(* IEC 61131-3 sources: volt/packages/volt-lsp-iec/test-corpus/pro2193/Device/Plc Logic/Application/09 Misc/Library Manager/L_IOM_IOModules, 22 files *)

(* ---- L_IOM_FAST_OUTP.dut ---- *)
TYPE L_IOM_FAST_OUTP :
STRUCT
	BYVALUE : BYTE;
	BYRUNNINGNUMBER : BYTE;
	WTIMETICK : WORD;
	DWTIMETICK : DWORD;
	XINUSE : BOOL;
END_STRUCT
END_TYPE

(* ---- L_IOM_FAST_OUTP_UNSORTED.dut ---- *)
TYPE L_IOM_FAST_OUTP_UNSORTED :
STRUCT
	BYDIGITALOUTPUTSEL : BYTE;
	BYVALUE : BYTE;
	WTIMETICK : WORD;
	DWTIMETICK : DWORD;
	XINUSE : BOOL;
END_STRUCT
END_TYPE

(* ---- L_IOM_FAST_RXTXPDO.dut ---- *)
TYPE L_IOM_FAST_RXTXPDO :
STRUCT
	WNUMBEROFEXCLUDES : WORD;
	WNUMBEROFENTRIES : WORD;
	WINDEX : WORD;
	BYFIXED : BYTE;
	BYMANDATORY : BYTE;
	WVIRTUAL : WORD;
	WSM : WORD;
	WSU : WORD;
	SNAME : STRING;
END_STRUCT
END_TYPE

(* ---- L_IOM_FAST_TXPDO.dut ---- *)
TYPE L_IOM_FAST_TXPDO :
STRUCT
	WINDEX : WORD;
	WSUBINDEX : WORD;
	WSIZE : WORD;
END_STRUCT
END_TYPE

(* ---- L_IOM_FASTIO_IO_ADDRESSES.dut ---- *)
TYPE L_IOM_FASTIO_IO_ADDRESSES :
STRUCT
	PBYVALUE : POINTER TO BYTE;
	PBYRUNNINGNUMBER : POINTER TO BYTE;
	PWTIMETICK : POINTER TO WORD;
END_STRUCT
END_TYPE

(* ---- L_IOM_FASTIO_OUT_STATE_INPUT.dut ---- *)
TYPE L_IOM_FASTIO_OUT_STATE_INPUT :
STRUCT
	PBYLASTRUNNINGNUMBER : POINTER TO BYTE;
	PBYNEXTRUNNINGNUMBER : POINTER TO BYTE;
	PBYSTATEFIFO : POINTER TO BYTE;
	PBYCOUNTFIFOENTRIES : POINTER TO BYTE;
	PDWABSOLUTECOUNTER : POINTER TO DWORD;
END_STRUCT
END_TYPE

(* ---- L_IOM_IEXTERNALTPINTERFACE.itf ---- *)
INTERFACE L_IOM_IEXTERNALTPINTERFACE
END_INTERFACE

METHOD CHECKABORTED : BOOL
VAR_INPUT
	TOUCHPROBECHANNEL : BYTE;
END_VAR
END_METHOD

METHOD CHECKCONFIGURATION : BOOL
VAR_INPUT
	TOUCHPROBESOURCE : BYTE;
	TOUCHPROBECHANNEL : BYTE;
	TOUCHPROBESIGNAL : BYTE;
	TOUCHPROBEEDGE : BYTE;
	TOUCHPROBEMODE : BYTE;
END_VAR
VAR_OUTPUT
	WERRORID : WORD := 0;
END_VAR
END_METHOD

METHOD CHECKNEWTP : BOOL
VAR_INPUT
	TOUCHPROBECHANNEL : BYTE;
	TOUCHPROBEEDGE : BYTE;
END_VAR
VAR_OUTPUT
	XTPPOSEDGE : BOOL;
	XTPNEGEDGE : BOOL;
	WTPTIMETICKPOSEDGE : WORD;
	WTPTIMETICKNEGEDGE : WORD;
	DWTPTIMETICKABSCOUNTER : DWORD;
END_VAR
END_METHOD

METHOD INITFORNEWTP : BOOL
VAR_INPUT
	TOUCHPROBECHANNEL : BYTE;
END_VAR
END_METHOD

METHOD SETABORT : BOOL
VAR_INPUT
	TOUCHPROBECHANNEL : BYTE;
END_VAR
END_METHOD

(* ---- CALCRXPDOOFFSETS131.pou ---- *)
FUNCTION CALCRXPDOOFFSETS131 : BOOL
VAR_INPUT
	PCONNECTOR : POINTER TO IoConfigConnector;
	WSLICEPOSITION : WORD;
	WPDOOFFSETBASE : WORD;
END_VAR
VAR_OUTPUT
	WPDOOFFSET : WORD;
	WPDONUMBEROFENTRIES : WORD;
END_VAR
END_FUNCTION

(* ---- CALCTXPDOOFFSETS131.pou ---- *)
FUNCTION CALCTXPDOOFFSETS131 : BOOL
VAR_INPUT
	PCONNECTOR : POINTER TO IoConfigConnector;
	WSLICEPOSITION : WORD;
	WPDOOFFSETBASE : WORD;
END_VAR
VAR_OUTPUT
	WPDOOFFSET : WORD;
	WPDONUMBEROFENTRIES : WORD;
END_VAR
END_FUNCTION

(* ---- FINDOWNSLICEPOSITIONS131.pou ---- *)
FUNCTION FINDOWNSLICEPOSITIONS131 : BOOL
VAR_INPUT
	M_HINTERFACE : POINTER TO IoConfigConnector;
	M_PCONNECTOR : POINTER TO IoConfigConnector;
	WMODULETYPE : WORD;
END_VAR
VAR_OUTPUT
	WSLICEPOSITION : WORD;
END_VAR
END_FUNCTION

(* ---- GETBOOLEANPROPERTY.pou ---- *)
FUNCTION GETBOOLEANPROPERTY : BOOL
VAR_INPUT
	STKEY : WSTRING;
END_VAR
END_FUNCTION

(* ---- GETCOMPANY.pou ---- *)
FUNCTION GETCOMPANY : WSTRING
END_FUNCTION

(* ---- GETNUMBERPROPERTY.pou ---- *)
FUNCTION GETNUMBERPROPERTY : DINT
VAR_INPUT
	STKEY : WSTRING;
END_VAR
END_FUNCTION

(* ---- GETTEXTPROPERTY.pou ---- *)
FUNCTION GETTEXTPROPERTY : WSTRING
VAR_INPUT
	STKEY : WSTRING;
END_VAR
END_FUNCTION

(* ---- GETTEXTPROPERTY2.pou ---- *)
FUNCTION GETTEXTPROPERTY2 : POINTER TO WSTRING
VAR_INPUT
	STKEY : WSTRING;
END_VAR
END_FUNCTION

(* ---- GETTITLE.pou ---- *)
FUNCTION GETTITLE : WSTRING
END_FUNCTION

(* ---- GETVERSION.pou ---- *)
FUNCTION GETVERSION : VERSION
END_FUNCTION

(* ---- GETVERSIONPROPERTY.pou ---- *)
FUNCTION GETVERSIONPROPERTY : VERSION
VAR_INPUT
	STKEY : WSTRING;
END_VAR
END_FUNCTION

(* ---- L_FASTIO_INREF.pou ---- *)
FUNCTION_BLOCK L_FASTIO_INREF EXTENDS IoDrvBase
VAR_INPUT
	XAABORTISACTIVE : ARRAY [0..3] OF BOOL;
END_VAR
VAR_OUTPUT
	IOVARIABLEADDRESSES : ARRAY [0..(FIFO_SIZE_MAX - 1)] OF L_IOM_FASTIO_IO_ADDRESSES;
	BYRISINGEDGEPARAMETERVALUE : BYTE;
	BYFALLINGEDGEPARAMETERVALUE : BYTE;
	BYMAXTPCOUNT : BYTE := 2;
	PDWABSOLUTECOUNTER : POINTER TO DWORD;
END_VAR
VAR
	CMPID_CMPLENZEFASTIO_INREF : DWORD := 16#1028200B;
	FIFO_SIZE_MAX : BYTE := 15;
	PARAM_ID_MODUL_IDENT : DWORD := 16#41000000;
	MODUL_IDENT_S207 : DWORD := 16#F0147C1;
	MODUL_IDENT_S208 : DWORD := 16#F0347C2;
	M_IIODRV : ICmpIoDrv;
	M_IIODRVPARAMETER : ICmpIoDrvParameter;
	XINPUTSVALID : BOOL := TRUE;
	XINPUTSVALIDACTCYCLE : BOOL := TRUE;
	XFIRSTEDGEDETECTED : BOOL := FALSE;
	ILASTRUNNINGNUMBER : ARRAY [1..4] OF INT := [-1, -1, -1, -1];
	BYNEWSIGNAL : ARRAY [1..4] OF BYTE := [0, 0, 0, 0];
	BYOLDSIGNAL : ARRAY [1..4] OF BYTE := [0, 0, 0, 0];
	FIFO_SIZE : BYTE;
	PMYFATHERCONNECT_68 : POINTER TO IoConfigConnector;
	PMYGRANDFATHERCONNECT_65 : POINTER TO IoConfigConnector;
	DWMODULIDENT : DWORD;
	PRESULT : POINTER TO SysTypes.RTS_IEC_RESULT;
	_XINITIALINPUTSTATEAVAILABLE : BOOL := FALSE;
	_ABYINITIALINPUTSTATE : ARRAY [0..1] OF BYTE;
	XFIRSTEDGETIMESTAMPVALID : BOOL := FALSE;
	DWFIRSTEDGETIMESTAMP : DWORD;
	BYINITIALINPUTSTATE : BYTE;
	FIRSTEDGEDETECTED : BOOL;
END_VAR
END_FUNCTION_BLOCK

METHOD INITIALIZE : UDINT
VAR_INPUT
	WMODULETYPE : UINT;
	DWINSTANCE : UDINT;
	PCONNECTOR : POINTER TO IoConfigConnector;
END_VAR
END_METHOD

METHOD FB_INIT : BOOL
VAR_INPUT
	BINITRETAINS : BOOL;
	BINCOPYCODE : BOOL;
END_VAR
END_METHOD

METHOD QUERYINTERFACE : POINTER TO POINTER TO BYTE
VAR_INPUT
	IID : DWORD;
	PRESULT : POINTER TO UDINT;
END_VAR
END_METHOD

METHOD IODRVUPDATECONFIGURATION : UDINT
VAR_INPUT
	PCONNECTORLIST : POINTER TO IoConfigConnector;
	NCOUNT : DINT;
END_VAR
END_METHOD

METHOD IODRVUPDATEMAPPING : UDINT
VAR_INPUT
	PTASKMAPLIST : POINTER TO IoConfigTaskMap;
	NCOUNT : DINT;
END_VAR
END_METHOD

METHOD IODRVGETCONNECTOR : POINTER TO IoConfigConnector
VAR_INPUT
	PRESULT : POINTER TO SysTypes.RTS_IEC_RESULT;
END_VAR
END_METHOD

METHOD CHECKABORTED : BOOL
VAR_INPUT
	TOUCHPROBECHANNEL : BYTE;
END_VAR
END_METHOD

METHOD CHECKCONFIGURATION : BOOL
VAR_INPUT
	TOUCHPROBESOURCE : BYTE;
	TOUCHPROBECHANNEL : BYTE;
	TOUCHPROBESIGNAL : BYTE;
	TOUCHPROBEEDGE : BYTE;
	TOUCHPROBEMODE : BYTE;
END_VAR
VAR_OUTPUT
	WERRORID : WORD := 0;
END_VAR
END_METHOD

METHOD CHECKNEWTP : BOOL
VAR_INPUT
	TOUCHPROBECHANNEL : BYTE;
	TOUCHPROBEEDGE : BYTE;
END_VAR
VAR_OUTPUT
	XTPPOSEDGE : BOOL;
	XTPNEGEDGE : BOOL;
	WTPTIMETICKPOSEDGE : WORD;
	WTPTIMETICKNEGEDGE : WORD;
	DWTPTIMETICKABSCOUNTER : DWORD;
END_VAR
END_METHOD

METHOD EDGEDETECTED : BOOL
VAR_INPUT
	TOUCHPROBEEDGE : BYTE;
	BYNEWSIGNAL : BYTE;
	BYOLDSIGNAL : BYTE;
	WTIMETICK : WORD;
END_VAR
VAR_OUTPUT
	XTPPOSEDGE : BOOL;
	XTPNEGEDGE : BOOL;
	WTPTIMETICKPOSEDGE : WORD;
	WTPTIMETICKNEGEDGE : WORD;
END_VAR
END_METHOD

METHOD INITFORNEWTP : BOOL
VAR_INPUT
	TOUCHPROBECHANNEL : BYTE;
END_VAR
END_METHOD

METHOD SETABORT : BOOL
VAR_INPUT
	TOUCHPROBECHANNEL : BYTE;
END_VAR
END_METHOD

(* ---- L_FASTIO_INREF_ECAT.pou ---- *)
FUNCTION_BLOCK L_FASTIO_INREF_ECAT EXTENDS L_FastIO_InRef
VAR
	WINITSTATE : WORD := 0;
	DWBUFFER : DWORD;
	L_ETC_COE_SDOWRITE1 : L_ETC_CoE_SdoWrite;
	L_ETC_GETMASTERSTATE1 : L_ETC_GetMasterState;
	WSLICEPOSITION : WORD;
	WPDOOFFSET : WORD;
	WPDONUMBEROFENTRIES : WORD;
	WECATSLAVEADR : WORD;
	PDWABSOLUTECOUNTERBPB : POINTER TO DWORD;
	PTASKMAPLISTFB : POINTER TO IoConfigTaskMap;
	PCONNECTORMAPFB : POINTER TO IoConfigConnectorMap;
	NCOUNTFB : DINT;
	ULIACTDCTIME_US : ULINT;
	ULIACTDCTIME_NS : ULINT;
	DWACTDCTIME_US : DWORD;
	WACTDCTIME_US : WORD;
END_VAR
END_FUNCTION_BLOCK

METHOD BEFOREREADINPUTS : INT
END_METHOD

METHOD FB_INIT : BOOL
VAR_INPUT
	BINITRETAINS : BOOL;
	BINCOPYCODE : BOOL;
END_VAR
END_METHOD

METHOD IODRVUPDATEMAPPING : UDINT
VAR_INPUT
	PTASKMAPLIST : POINTER TO IoConfigTaskMap;
	NCOUNT : DINT;
END_VAR
END_METHOD

(* ---- L_FASTIO_OUTREF.pou ---- *)
FUNCTION_BLOCK L_FASTIO_OUTREF EXTENDS IoDrvBase
VAR_OUTPUT
	INPUTVARIABLEADDRESSES : L_IOM_FASTIO_OUT_STATE_INPUT;
	FIFOVARIABLEADDRESSES : ARRAY [0..(FIFO_SIZE_MAX - 1)] OF L_IOM_FASTIO_IO_ADDRESSES;
END_VAR
VAR
	CMPID_CMPLENZEFASTIO_OUTREF : DWORD := 16#1028200C;
	FIFO_SIZE_MAX : BYTE := 15;
	PARAM_ID_MODUL_IDENT : DWORD := 16#41000000;
	MODUL_IDENT_S310 : DWORD := 16#F4157E1;
	MODUL_IDENT_S311 : DWORD := 16#F4357E2;
	M_IIODRV : ICmpIoDrv;
	M_IIODRVPARAMETER : ICmpIoDrvParameter;
	M_BYNEXTFIFOINDEX : BYTE;
	M_BYLASTOUTPUTVALUE : BYTE := 16#30;
	M_BYLASTRUNNINGNUMBER : BYTE;
	M_DWMIKROSECTICKLAST : DWORD;
	M_IMIKROSECTICKCYCLECOUNT : INT;
	AFIFOUNSORTED : ARRAY [0..7] OF L_IOM_FAST_OUTP_UNSORTED;
	M_BYNEXTFIFOUNSORTEDINDEX : BYTE;
	FIFO_SIZE : BYTE := 8;
	BYMAXOUTPCOUNT : BYTE := 2;
	PMYFATHERCONNECT_68 : POINTER TO IoConfigConnector;
	PMYGRANDFATHERCONNECT_65 : POINTER TO IoConfigConnector;
	DWMODULIDENT : DWORD;
	PRESULT : POINTER TO SysTypes.RTS_IEC_RESULT;
	PIOCONFIGPARAMETER : POINTER TO IoConfigParameter;
END_VAR
END_FUNCTION_BLOCK

METHOD AFTERWRITEOUTPUTS : INT
END_METHOD

METHOD BEFOREWRITEOUTPUTS : INT
END_METHOD

METHOD INITIALIZE : UDINT
VAR_INPUT
	WMODULETYPE : UINT;
	DWINSTANCE : UDINT;
	PCONNECTOR : POINTER TO IoConfigConnector;
END_VAR
END_METHOD

METHOD INSERTNEWFIFOENTRY : INT
VAR_INPUT
	BYDIGITALOUTPUTSEL : BYTE;
	BYVALUE : BYTE;
	WTIMERTICK : WORD;
END_VAR
END_METHOD

METHOD INSERTNEWFIFOENTRYINTERN : INT
VAR_INPUT
	BYDIGITALOUTPUTSEL : BYTE;
	BYVALUE : BYTE;
	WTIMERTICK : WORD;
END_VAR
END_METHOD

METHOD FB_INIT : BOOL
VAR_INPUT
	BINITRETAINS : BOOL;
	BINCOPYCODE : BOOL;
END_VAR
END_METHOD

METHOD QUERYINTERFACE : POINTER TO POINTER TO BYTE
VAR_INPUT
	IID : DWORD;
	PRESULT : POINTER TO UDINT;
END_VAR
END_METHOD

METHOD IODRVUPDATECONFIGURATION : UDINT
VAR_INPUT
	PCONNECTORLIST : POINTER TO IoConfigConnector;
	NCOUNT : DINT;
END_VAR
END_METHOD

METHOD IODRVUPDATEMAPPING : UDINT
VAR_INPUT
	PTASKMAPLIST : POINTER TO IoConfigTaskMap;
	NCOUNT : DINT;
END_VAR
END_METHOD

METHOD IODRVGETCONNECTOR : POINTER TO IoConfigConnector
VAR_INPUT
	PRESULT : POINTER TO SysTypes.RTS_IEC_RESULT;
END_VAR
END_METHOD

(* ---- L_FASTIO_OUTREF_ECAT.pou ---- *)
FUNCTION_BLOCK L_FASTIO_OUTREF_ECAT EXTENDS L_FastIO_OutRef
VAR
	WSLICEPOSITION : WORD;
	WPDOOFFSET : WORD;
	WPDONUMBEROFENTRIES : WORD;
	L_ETC_GETMASTERSTATE1 : L_ETC_GetMasterState;
	PTASKMAPLISTFB : POINTER TO IoConfigTaskMap;
	PCONNECTORMAPFB : POINTER TO IoConfigConnectorMap;
	PCONNECTORLISTFB : POINTER TO IoConfigConnector;
	NCOUNTFB : DINT;
	PDWABSOLUTECOUNTERBPB : POINTER TO DWORD;
	ULIACTDCTIME_US : ULINT;
	ULIACTDCTIME_NS : ULINT;
	DWACTDCTIME_NS : DWORD;
	DWACTDCTIME_US : DWORD;
	WACTDCTIME_US : WORD;
	WINITSTATE : WORD;
END_VAR
END_FUNCTION_BLOCK

METHOD BEFOREREADINPUTS : INT
END_METHOD

METHOD FB_INIT : BOOL
VAR_INPUT
	BINITRETAINS : BOOL;
	BINCOPYCODE : BOOL;
END_VAR
END_METHOD

METHOD IODRVUPDATEMAPPING : UDINT
VAR_INPUT
	PTASKMAPLIST : POINTER TO IoConfigTaskMap;
	NCOUNT : DINT;
END_VAR
END_METHOD
